Fanuc KAREL source: kb00131.KL

-- PROVISIONAL review KL for V940-1; original PC SHA256 8dc4f2719635d0bf885a47122d0144157f93e40ae201861b4818737d5e6a108a
-- Incomplete behavior may be omitted. Consult companion uncertainty JSON. Do not deploy.
PROGRAM KB00131
%NOLOCKGROUP
BEGIN
  -- V9_ZERO_TABLE_METADATA_HINT layout=0002_ascii; no indexed target words; source/name/runtime held
  -- UNRESOLVED_PC offsets 5-14; opcodes 3F,75
  -- UNRESOLVED_PC offsets 19-26; opcodes 9D,23
  -- UNRESOLVED_PC offsets 31-38; opcodes 9D,23
  -- UNRESOLVED_PC offsets 43-50; opcodes 9D,23
  -- UNRESOLVED_PC offsets 55-64; opcodes 3F,75
  -- UNRESOLVED_PC offsets 69-76; opcodes 9D,23
  -- UNRESOLVED_PC offsets 81-88; opcodes 9D,23
  -- UNRESOLVED_PC offsets 93-143; opcodes 27,22,2A,22,22,22,22,2A,22,22,31
  -- UNRESOLVED_PC offsets 148-152; opcodes 7F
END KB00131
